(* CODESYS project Overview_current.export

Project tree, tasks and I/O mapping:
  visualisation Overview
*)

// /Overview
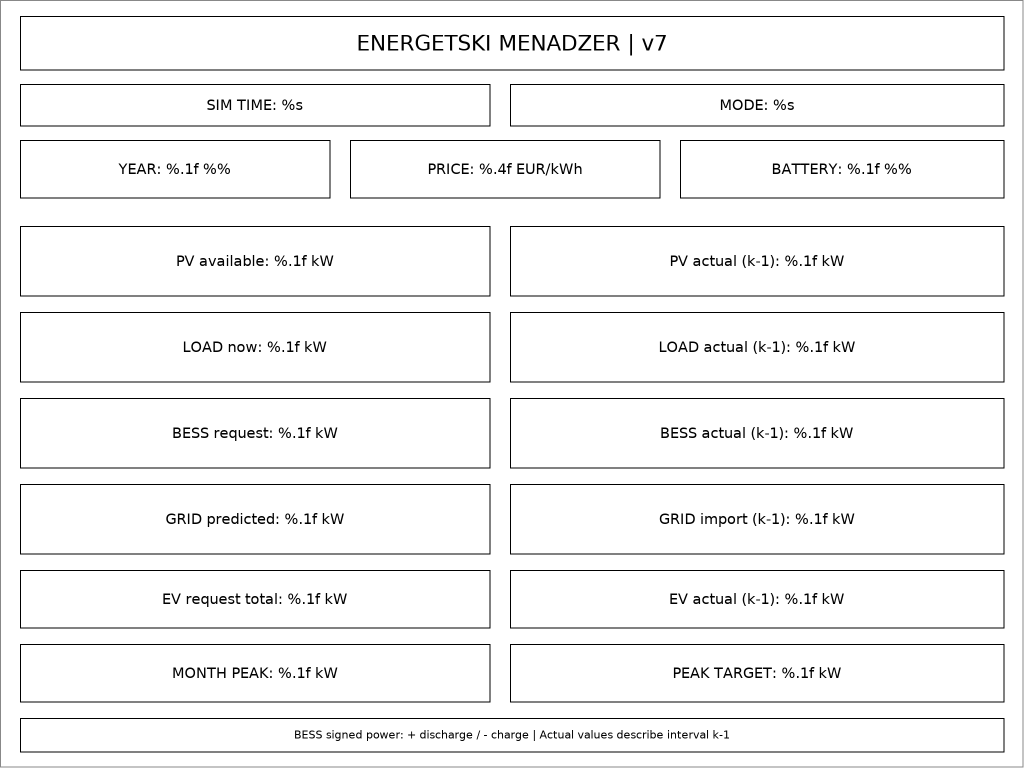
VISUALIZATION Overview  // 1024x768
    Rectangle (20,16 984x54), "ENERGETSKI MENADZER | v7"
    Rectangle (20,84 470x42), "SIM TIME: %s", text variable: Team_HMI.sDateTime
    Rectangle (510,84 494x42), "MODE: %s", text variable: Team_HMI.sPriceMode
    Rectangle (20,140 310x58), "YEAR: %.1f %%", text variable: Team_HMI.rProgressPct
    Rectangle (350,140 310x58), "PRICE: %.4f EUR/kWh", text variable: Team_HMI.rPrice
    Rectangle (680,140 324x58), "BATTERY: %.1f %%", text variable: Team_HMI.rSoc
    Rectangle (20,226 470x70), "PV available: %.1f kW", text variable: Team_HMI.rFneAvail
    Rectangle (510,226 494x70), "PV actual (k-1): %.1f kW", text variable: Team_HMI.rFneAct
    Rectangle (20,312 470x70), "LOAD now: %.1f kW", text variable: Team_HMI.rFec
    Rectangle (510,312 494x70), "LOAD actual (k-1): %.1f kW", text variable: Team_HMI.rFecPrev
    Rectangle (20,398 470x70), "BESS request: %.1f kW", text variable: Team_HMI.rBessReq
    Rectangle (510,398 494x70), "BESS actual (k-1): %.1f kW", text variable: Team_HMI.rBessAct
    Rectangle (20,484 470x70), "GRID predicted: %.1f kW", text variable: Team_HMI.rGridPred
    Rectangle (510,484 494x70), "GRID import (k-1): %.1f kW", text variable: Team_HMI.rImportAct
    Rectangle (20,570 470x58), "EV request total: %.1f kW", text variable: Team_HMI.rEvReqSum
    Rectangle (510,570 494x58), "EV actual (k-1): %.1f kW", text variable: Team_HMI.rEvActSum
    Rectangle (20,644 470x58), "MONTH PEAK: %.1f kW", text variable: Team_HMI.rPeakMonth
    Rectangle (510,644 494x58), "PEAK TARGET: %.1f kW", text variable: Team_HMI.rPeakTarget
    Rectangle (20,718 984x34), "BESS signed power: + discharge / - charge | Actual values describe interval k-1"
END_VISUALIZATION
